(* IEC 61131-3 sources: ZPLC/conformance/harness, 3 files *)

(* ---- vf-001-bool-output-toggles.st ---- *)
PROGRAM Toggle
VAR
  q AT %QX0.0 : BOOL;
END_VAR
  q := NOT q;
END_PROGRAM

(* ---- vf-001-input-reaches-output.st ---- *)
PROGRAM Copy
VAR
  go AT %IX0.0 : BOOL;
  lamp AT %QX0.0 : BOOL;
END_VAR
  lamp := go;
END_PROGRAM

(* ---- vf-001-vm-fault-is-observed.st ---- *)
PROGRAM Fault
VAR
  zero : INT;
  quotient AT %QW0 : INT;
END_VAR
  quotient := 100 / zero;
END_PROGRAM
